Fanuc KAREL source: KC00035.KL

PROGRAM KC00035
%NOLOCKGROUP
VAR
  I: INTEGER
  J: INTEGER
  K: INTEGER
  R: REAL
  B: BOOLEAN
  S: STRING[80]
  T: STRING[80]
  P: PATH
  Q: PATH
  AI: ARRAY[8] OF INTEGER
  AB: ARRAY[244] OF BYTE
  F: FILE
BEGIN
  XML_SCAN(F,S,I,J,K)
END KC00035
